// TIA Portal V20 export
VAR_GLOBAL   // PLC tag table "T2_Variables"
   T2_M_Falso AT %M950.0 : Bool;   // Prueba IA 2: siempre FALSE (nadie la escribe)
   T2_MW_Prueba AT %MW952 : Int;   // Prueba IA 2: palabra de marcas
END_VAR
